(*
    What FB_PneumaticActuator and FB_MPA share: the position state from the two limit switches,
    and the timeout of an output that does not reach its limit switch.
*)
INTERFACE I_PneumaticCore

PROPERTY State : E_PnuematicActuatorPositionState
GET
END_GET
END_PROPERTY

PROPERTY InsertTimedOut : BOOL
GET
END_GET
END_PROPERTY

PROPERTY RetractTimedOut : BOOL
GET
END_GET
END_PROPERTY

PROPERTY InsertTimeoutElapsed : BOOL
GET
END_GET
END_PROPERTY

PROPERTY RetractTimeoutElapsed : BOOL
GET
END_GET
END_PROPERTY

END_INTERFACE

(* stored: Version 1.1.0.1
   Itf I_PneumaticCore: Id {ffa8e96f-fadc-4004-a845-6738863ddf56}
   Property State: Id {05fc219d-f37b-4cfd-98a7-0424a2548a3d}
   Get Get: Id {6e1f9b34-27a8-4d5c-b0e3-8a7c2d9f1b46}
   Property InsertTimedOut: Id {c8e41a07-6d2b-4f93-a5b0-3e97d1f60c28}
   Get Get: Id {51f0b9d3-7a84-4c6e-b2d5-0e8a3c971f46}
   Property RetractTimedOut: Id {2f6d83b1-94e0-4a7c-8d15-b7c3e0a92f64}
   Get Get: Id {9b04e7c5-1d38-4f2a-a6c9-84e1f5b03d72}
   Property InsertTimeoutElapsed: Id {5941fd68-877e-4429-bc96-49fae16c8b15}
   Get Get: Id {82cadbff-b216-4255-a475-ece2e199a942}
   Property RetractTimeoutElapsed: Id {a5ee096b-328a-4318-9ae0-00a4c6ca1216}
   Get Get: Id {94d624cb-6114-44e3-99ac-1ca3de2e759e} *)
